// // MIGRATION DRAFT: not included in PLC compilation.
// // Reference: Reference_Project/Screens.scl, object OT_Charge_Commands.
// // Types, globals, calls, units and behavior require manual reconciliation.
// // See docs/TIA_Missing_Blocks.md before importing as PLC code.
FUNCTION OT_Charge_Commands : BOOL
// 
//    VAR_IN_OUT
//       Auto_Test : Auto_Test;
//    END_VAR

// // MIGRATION DRAFT: not included in PLC compilation.
// // Reference: Reference_Project/Screens.scl, object OT_Charge_Commands.
// // Types, globals, calls, units and behavior require manual reconciliation.
// // See docs/TIA_Missing_Blocks.md before importing as PLC code.
// OrderTable_HMI.Manual_order := Auto_Test.Manual;
// 
// 	IF Auto_Test.Pallet_Type = 'C' THEN
// 	    OrderTable_HMI.Pallet_Type := 1;
// 	ELSIF Auto_Test.Pallet_Type = 'E' THEN
// 	    OrderTable_HMI.Pallet_Type := 2;
// 	END_IF;
// 
// 	IF Auto_Test.Tower_1_Pallet_Alignment = 'R' THEN
// 	    OrderTable_HMI.Tower_1_Pallet_Alignment := 1;
// 	ELSIF Auto_Test.Tower_1_Pallet_Alignment = 'L' THEN
// 	    OrderTable_HMI.Tower_1_Pallet_Alignment := 2;
// 	END_IF;
// 
// 	IF Auto_Test.Tower_2_Pallet_Alignment = 'R' THEN
// 	    OrderTable_HMI.Tower_2_Pallet_Alignment := 1;
// 	ELSIF Auto_Test.Tower_2_Pallet_Alignment = 'L' THEN
// 	    OrderTable_HMI.Tower_2_Pallet_Alignment := 2;
// 	END_IF;
// 
// 	IF Auto_Test.Extractor_Pallet_Alignment = 'R' THEN
// 	    OrderTable_HMI.Extractor_Pallet_Alignment := 1;
// 	ELSIF Auto_Test.Extractor_Pallet_Alignment = 'L' THEN
// 	    OrderTable_HMI.Extractor_Pallet_Alignment := 2;
// 	ELSIF Auto_Test.Extractor_Pallet_Alignment = 'C' THEN
// 	    OrderTable_HMI.Extractor_Pallet_Alignment := 3;
// 	END_IF;
// 	OrderTable_HMI.From_level := Auto_Test.From_level;
// 	OrderTable_HMI.To_level := Auto_Test.To_level;
// 	OrderTable_HMI.Testing_Time := Auto_Test.Testing_Time;
// 	OrderTable_HMI.Numer_of_cycles := Auto_Test.Numer_of_cycles;
// 	OrderTable_HMI.Level := UINT_TO_BYTE(Auto_Test.Level);
// 	OrderTable_HMI.Tower := UINT_TO_BYTE(Auto_Test.Tower);

END_FUNCTION

(* stored: Version 1.1.0.1
   POU OT_Charge_Commands: Id {99cc0188-a0a3-500c-a760-8d20debe74d7}, SpecialFunc None *)
